Staubli VAL3: initArmInfo.pgx

program initArmInfo()
  local string l_sLanguage
  local string l_sMounting
begin
  //*******************************************************
  db:utLbl_Axis_Data.Common.sText="4axis"
  //*******************************************************
  //Get mounting property
  //*******************************************************
  l_sMounting=getVersion("Arm Mounting")
  switch l_sMounting
    case "floor"
      db:sMounting="Floor"
      db:utCbx_Mounting_Data.Common.sValue="Floor"
    break
    case "ceiling"
      db:sMounting="Ceiling"
      db:utCbx_Mounting_Data.Common.sValue="Ceiling"
    break
    default
      db:sMounting="Null"
      db:utCbx_Mounting_Data.Common.sValue=""
    break
  endSwitch
  //*******************************************************
  //Get system language
  //*******************************************************
  l_sLanguage=getLanguage()
  switch l_sLanguage
    case "chinese"
      db:sLanguage="chinese"
      db:utCbx_Language_Data.Common.sValue="Chinese"
    break
    case "english"
      db:sLanguage="english"
      db:utCbx_Language_Data.Common.sValue="English"
    break
    default
      db:sLanguage="english"
      db:utCbx_Language_Data.Common.sValue="English"
    break
  endSwitch
  //
  //*******************************************************
  //Initialize the flange as the current tool
  //*******************************************************
  call db:updateTool(0,false)
end
